// TIA Portal V21 export
// export: Created 2026-08-21T20:18:51.3701793Z, ExportSetting None, DisplayName Totally Integrated Automation Portal, DisplayVersion V21, DisplayName STEP 7 Professional, DisplayVersion V21, DisplayName STEP 7 Safety, DisplayVersion V21, DisplayName Tech WebApplication, DisplayVersion V21, DisplayName WinCC Basic/Comfort/Advanced, DisplayVersion V21, DisplayName WinCC Professional, DisplayVersion V21, DisplayName WinCC Unified, DisplayVersion V21
ORGANIZATION_BLOCK "Startup"   // OB100, FBD, Startup
TITLE = "Complete Restart"
{ S7_Optimized_Access := 'TRUE' }
// stored: SetENOAutomatically false
   VAR_INPUT
      LostRetentive : Bool;   // True if retentive data are lost
      LostRTC : Bool;   // True if date and time are lost
   END_VAR
BEGIN

REGION Network 1
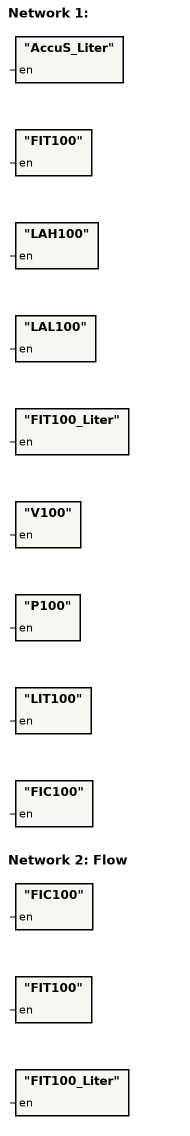
   "AccuS_Liter"();
   "FIT100"();
   "LAH100"();
   "LAL100"();
   "FIT100_Liter"();
   "V100"();
   "P100"();
   "LIT100"();
   "FIC100"();
END_REGION

REGION Network 2: Flow
   "FIC100"();
   "FIT100"();
   "FIT100_Liter"();
END_REGION

REGION Network 3: Level
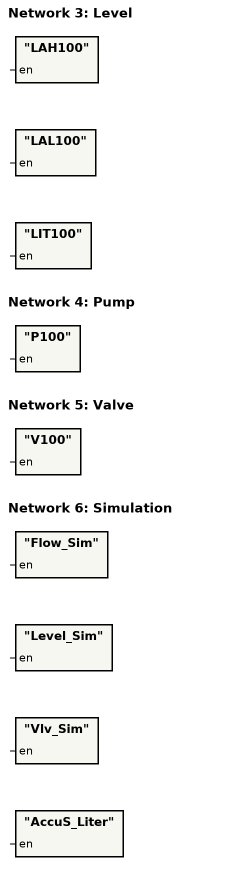
   "LAH100"();
   "LAL100"();
   "LIT100"();
END_REGION

REGION Network 4: Pump
   "P100"();
END_REGION

REGION Network 5: Valve
   "V100"();
END_REGION

REGION Network 6: Simulation
   "Flow_Sim"();
   "Level_Sim"();
   "Vlv_Sim"();
   "AccuS_Liter"();
END_REGION
END_ORGANIZATION_BLOCK
